// TIA Portal V20 export
// export: Created 2026-10-19T18:06:12.0545381Z, ExportSetting WithDefaults, DisplayName Totally Integrated Automation Portal, DisplayVersion V20 Update 6, DisplayName TIA Portal Openness, DisplayVersion V20 Update 6, DisplayName TIA Portal Version Control Interface, DisplayVersion V20 Update 6, DisplayName SINAMICS Startdrive Advanced, DisplayVersion V20 SP1, DisplayName SINAMICS Startdrive G130, G150, S120, S150, SINAMICS MV, G220, S200, S210, DisplayVersion V20 SP1, DisplayName SINAMICS Startdrive G110M, G120, G120C, G120D, G120P, G115D, DisplayVersion V20 SP1, DisplayName STEP 7 Professional, DisplayVersion V20 Update 6, DisplayName STEP 7 Safety, DisplayVersion V20 Update 2, DisplayName WinCC Basic/Comfort/Advanced, DisplayVersion V20 Update 6, DisplayName WinCC Unified, DisplayVersion V20 Update 6
FUNCTION "MT_ACT_Application" : Void   // FC30, LAD
{ S7_Optimized_Access := 'FALSE' }
VERSION : 0.1
// stored: AutoNumber true, IsIECCheckEnabled false, SetENOAutomatically false, UDAEnableTagReadback false
BEGIN

REGION Network 1: Cyclic Weighing Data
   // All the cyclical read and write commands can be issued from this Function Block.
   // The cyclic commands are triggered following a positive trigger. These commands are Tare Immediate, Tare Stable, Zero Immediate, Zero Stable, Pretare and Clear Tare. 
   // Upon successful execution of these commands, the DONE output bit will be set ON.
   // ERROR output bit will be set on if there is an error with the command execution.
   // Note: Only one cyclic command is possible at any one time.
   // If Net weight is required after executed a zero or tare command, insert decimal value "3" into the "WeightCmd" variable before triggering the cyclic scale command. Else, with decimal value "1" in the "WeightCmd" variable, the Function Block will return Gross Weight after the cyclic scale command. 
   // "DataOK" bit is set ON when the scale is in operation mode, not overloaded and not underload.
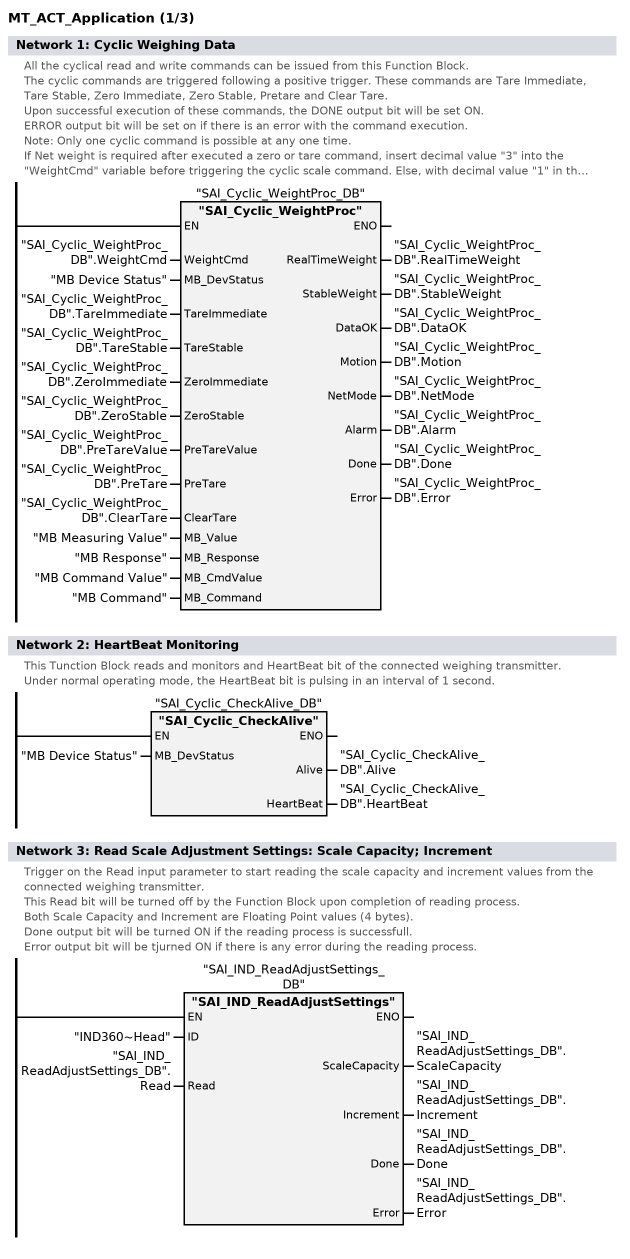
   RUNG wire#powerrail
      "SAI_Cyclic_WeightProc_DB"(WeightCmd := "SAI_Cyclic_WeightProc_DB".WeightCmd, MB_DevStatus := "MB Device Status", TareImmediate := "SAI_Cyclic_WeightProc_DB".TareImmediate, TareStable := "SAI_Cyclic_WeightProc_DB".TareStable, ZeroImmediate := "SAI_Cyclic_WeightProc_DB".ZeroImmediate, ZeroStable := "SAI_Cyclic_WeightProc_DB".ZeroStable, PreTareValue := "SAI_Cyclic_WeightProc_DB".PreTareValue, PreTare := "SAI_Cyclic_WeightProc_DB".PreTare, ClearTare := "SAI_Cyclic_WeightProc_DB".ClearTare, MB_Value := "MB Measuring Value", MB_Response := "MB Response", MB_CmdValue := "MB Command Value", MB_Command := "MB Command", RealTimeWeight => "SAI_Cyclic_WeightProc_DB".RealTimeWeight, StableWeight => "SAI_Cyclic_WeightProc_DB".StableWeight, DataOK => "SAI_Cyclic_WeightProc_DB".DataOK, Motion => "SAI_Cyclic_WeightProc_DB".Motion, NetMode => "SAI_Cyclic_WeightProc_DB".NetMode, Alarm => "SAI_Cyclic_WeightProc_DB".Alarm, Done => "SAI_Cyclic_WeightProc_DB".Done, Error => "SAI_Cyclic_WeightProc_DB".Error)
   END_RUNG
   // the same network as SCL:
   "SAI_Cyclic_WeightProc_DB"(WeightCmd := "SAI_Cyclic_WeightProc_DB".WeightCmd,   // "SAI_Cyclic_WeightProc"
                           MB_DevStatus := "MB Device Status",
                           TareImmediate := "SAI_Cyclic_WeightProc_DB".TareImmediate,
                           TareStable := "SAI_Cyclic_WeightProc_DB".TareStable,
                           ZeroImmediate := "SAI_Cyclic_WeightProc_DB".ZeroImmediate,
                           ZeroStable := "SAI_Cyclic_WeightProc_DB".ZeroStable,
                           PreTareValue := "SAI_Cyclic_WeightProc_DB".PreTareValue,
                           PreTare := "SAI_Cyclic_WeightProc_DB".PreTare,
                           ClearTare := "SAI_Cyclic_WeightProc_DB".ClearTare,
                           MB_Value := "MB Measuring Value",
                           MB_Response := "MB Response",
                           MB_CmdValue := "MB Command Value",
                           MB_Command := "MB Command",
                           RealTimeWeight => "SAI_Cyclic_WeightProc_DB".RealTimeWeight,
                           StableWeight => "SAI_Cyclic_WeightProc_DB".StableWeight,
                           DataOK => "SAI_Cyclic_WeightProc_DB".DataOK,
                           Motion => "SAI_Cyclic_WeightProc_DB".Motion,
                           NetMode => "SAI_Cyclic_WeightProc_DB".NetMode,
                           Alarm => "SAI_Cyclic_WeightProc_DB".Alarm,
                           Done => "SAI_Cyclic_WeightProc_DB".Done,
                           Error => "SAI_Cyclic_WeightProc_DB".Error);
END_REGION

REGION Network 2: HeartBeat Monitoring
   // This Tunction Block reads and monitors and HeartBeat bit of the connected weighing transmitter.
   // Under normal operating mode, the HeartBeat bit is pulsing in an interval of 1 second.
   RUNG wire#powerrail
      "SAI_Cyclic_CheckAlive_DB"(MB_DevStatus := "MB Device Status", Alive => "SAI_Cyclic_CheckAlive_DB".Alive, HeartBeat => "SAI_Cyclic_CheckAlive_DB".HeartBeat)
   END_RUNG
   // the same network as SCL:
   "SAI_Cyclic_CheckAlive_DB"(MB_DevStatus := "MB Device Status",   // "SAI_Cyclic_CheckAlive"
                           Alive => "SAI_Cyclic_CheckAlive_DB".Alive,
                           HeartBeat => "SAI_Cyclic_CheckAlive_DB".HeartBeat);
END_REGION

REGION Network 3: Read Scale Adjustment Settings: Scale Capacity; Increment
   // Trigger on the Read input parameter to start reading the scale capacity and increment values from the connected weighing transmitter.
   // This Read bit will be turned off by the Function Block upon completion of reading process.
   // Both Scale Capacity and Increment are Floating Point values (4 bytes).
   // Done output bit will be turned ON if the reading process is successfull.
   // Error output bit will be tjurned ON if there is any error during the reading process.
   RUNG wire#powerrail
      "SAI_IND_ReadAdjustSettings_DB"(ID := "IND360~Head", Read := "SAI_IND_ReadAdjustSettings_DB".Read, ScaleCapacity => "SAI_IND_ReadAdjustSettings_DB".ScaleCapacity, Increment => "SAI_IND_ReadAdjustSettings_DB".Increment, Done => "SAI_IND_ReadAdjustSettings_DB".Done, Error => "SAI_IND_ReadAdjustSettings_DB".Error)
   END_RUNG
   // the same network as SCL:
   "SAI_IND_ReadAdjustSettings_DB"(ID := "IND360~Head",   // "SAI_IND_ReadAdjustSettings"
                           Read := "SAI_IND_ReadAdjustSettings_DB".Read,
                           ScaleCapacity => "SAI_IND_ReadAdjustSettings_DB".ScaleCapacity,
                           Increment => "SAI_IND_ReadAdjustSettings_DB".Increment,
                           Done => "SAI_IND_ReadAdjustSettings_DB".Done,
                           Error => "SAI_IND_ReadAdjustSettings_DB".Error);
END_REGION

REGION Network 4: Write new Scale Adjustment Settings: Scale Capacity; Increment
   // Trigger on the Write input parameter to start writing the new scale capacity and increment settings to the connected weighing transmitter.
   // Both Scale Capacity and Increment are Floating Point values (4 bytes).
   // Make sure both settings are valid and correct before triggering the Write input bit.
   // This Write bit will be turned off by the Function Block upon completion of writing process.
   // Done output bit will be set ON if the reading process is successfull.
   // Error output bit will be set ON if there is any error during the reading process.
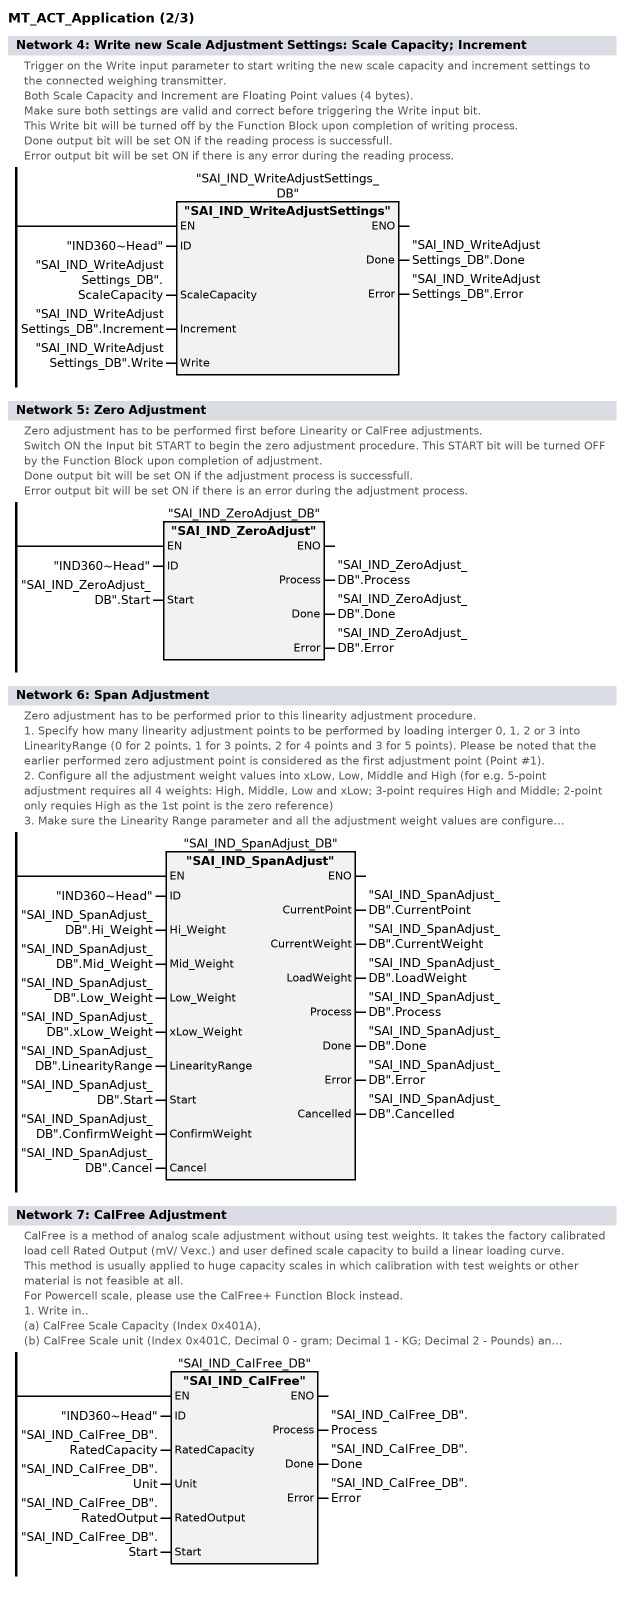
   RUNG wire#powerrail
      "SAI_IND_WriteAdjustSettings_DB"(ID := "IND360~Head", ScaleCapacity := "SAI_IND_WriteAdjustSettings_DB".ScaleCapacity, Increment := "SAI_IND_WriteAdjustSettings_DB".Increment, Write := "SAI_IND_WriteAdjustSettings_DB".Write, Done => "SAI_IND_WriteAdjustSettings_DB".Done, Error => "SAI_IND_WriteAdjustSettings_DB".Error)
   END_RUNG
   // the same network as SCL:
   "SAI_IND_WriteAdjustSettings_DB"(ID := "IND360~Head",   // "SAI_IND_WriteAdjustSettings"
                           ScaleCapacity := "SAI_IND_WriteAdjustSettings_DB".ScaleCapacity,
                           Increment := "SAI_IND_WriteAdjustSettings_DB".Increment,
                           Write := "SAI_IND_WriteAdjustSettings_DB".Write,
                           Done => "SAI_IND_WriteAdjustSettings_DB".Done,
                           Error => "SAI_IND_WriteAdjustSettings_DB".Error);
END_REGION

REGION Network 5: Zero Adjustment
   // Zero adjustment has to be performed first before Linearity or CalFree adjustments.
   // Switch ON the Input bit START to begin the zero adjustment procedure. This START bit will be turned OFF by the Function Block upon completion of adjustment. 
   // Done output bit will be set ON if the adjustment process is successfull.
   // Error output bit will be set ON if there is an error during the adjustment process.
   RUNG wire#powerrail
      "SAI_IND_ZeroAdjust_DB"(ID := "IND360~Head", Start := "SAI_IND_ZeroAdjust_DB".Start, Process => "SAI_IND_ZeroAdjust_DB".Process, Done => "SAI_IND_ZeroAdjust_DB".Done, Error => "SAI_IND_ZeroAdjust_DB".Error)
   END_RUNG
   // the same network as SCL:
   "SAI_IND_ZeroAdjust_DB"(ID := "IND360~Head",   // "SAI_IND_ZeroAdjust"
                           Start := "SAI_IND_ZeroAdjust_DB".Start,
                           Process => "SAI_IND_ZeroAdjust_DB".Process,
                           Done => "SAI_IND_ZeroAdjust_DB".Done,
                           Error => "SAI_IND_ZeroAdjust_DB".Error);
END_REGION

REGION Network 6: Span Adjustment
   // Zero adjustment has to be performed prior to this linearity adjustment procedure.
   // 
   // 1. Specify how many linearity adjustment points to be performed by loading interger 0, 1, 2 or 3 into LinearityRange (0 for 2 points, 1 for 3 points, 2 for 4 points and 3 for 5 points). Please be noted that the earlier performed zero adjustment point is considered as the first adjustment point (Point #1).
   // 
   // 2. Configure all the adjustment weight values into xLow, Low, Middle and High (for e.g. 5-point adjustment requires all 4 weights: High, Middle, Low and xLow; 3-point requires High and Middle; 2-point only requies High as the 1st point is the zero reference)
   // 
   // 3. Make sure the Linearity Range parameter and all the adjustment weight values are configured correctly before starting the adjustment process. Invalid or incomplete parameters will cause the Function Block to turn on the Error output bit.
   // 
   // 4. Trigger ON  Input Start bit to start the span adjustment. This Start bit will be turned off by the Function Block upon completion/ cancellation or error condition. 
   // 
   // 5. Once started, CurrentPoint shows the current linearity point to be adjusted; CurrentWeight shows current adjustment weight to be loaded onto the scale. The LoadWeight output bit will be set ON to request for new adjustment weight. 
   // 
   // 6. After loading the new adjustment weight, acknowledge this by triggering the ConfirmWeight parameter (boolean) ON. The Function Block will then proceed to the next adjustment point and turn off this ConfirmWeight bit.
   // 
   // 7. Output bit - Process signifies that the adjustment of current point is in process.
   // 
   // 8. Input Parameter Bit Cancel is used to cancel/ abort the adjustment process
   RUNG wire#powerrail
      "SAI_IND_SpanAdjust_DB"(ID := "IND360~Head", Hi_Weight := "SAI_IND_SpanAdjust_DB".Hi_Weight, Mid_Weight := "SAI_IND_SpanAdjust_DB".Mid_Weight, Low_Weight := "SAI_IND_SpanAdjust_DB".Low_Weight, xLow_Weight := "SAI_IND_SpanAdjust_DB".xLow_Weight, LinearityRange := "SAI_IND_SpanAdjust_DB".LinearityRange, Start := "SAI_IND_SpanAdjust_DB".Start, ConfirmWeight := "SAI_IND_SpanAdjust_DB".ConfirmWeight, Cancel := "SAI_IND_SpanAdjust_DB".Cancel, CurrentPoint => "SAI_IND_SpanAdjust_DB".CurrentPoint, CurrentWeight => "SAI_IND_SpanAdjust_DB".CurrentWeight, LoadWeight => "SAI_IND_SpanAdjust_DB".LoadWeight, Process => "SAI_IND_SpanAdjust_DB".Process, Done => "SAI_IND_SpanAdjust_DB".Done, Error => "SAI_IND_SpanAdjust_DB".Error, Cancelled => "SAI_IND_SpanAdjust_DB".Cancelled)
   END_RUNG
   // the same network as SCL:
   "SAI_IND_SpanAdjust_DB"(ID := "IND360~Head",   // "SAI_IND_SpanAdjust"
                           Hi_Weight := "SAI_IND_SpanAdjust_DB".Hi_Weight,
                           Mid_Weight := "SAI_IND_SpanAdjust_DB".Mid_Weight,
                           Low_Weight := "SAI_IND_SpanAdjust_DB".Low_Weight,
                           xLow_Weight := "SAI_IND_SpanAdjust_DB".xLow_Weight,
                           LinearityRange := "SAI_IND_SpanAdjust_DB".LinearityRange,
                           Start := "SAI_IND_SpanAdjust_DB".Start,
                           ConfirmWeight := "SAI_IND_SpanAdjust_DB".ConfirmWeight,
                           Cancel := "SAI_IND_SpanAdjust_DB".Cancel,
                           CurrentPoint => "SAI_IND_SpanAdjust_DB".CurrentPoint,
                           CurrentWeight => "SAI_IND_SpanAdjust_DB".CurrentWeight,
                           LoadWeight => "SAI_IND_SpanAdjust_DB".LoadWeight,
                           Process => "SAI_IND_SpanAdjust_DB".Process,
                           Done => "SAI_IND_SpanAdjust_DB".Done,
                           Error => "SAI_IND_SpanAdjust_DB".Error,
                           Cancelled => "SAI_IND_SpanAdjust_DB".Cancelled);
END_REGION

REGION Network 7: CalFree Adjustment
   // CalFree is a method of analog scale adjustment without using test weights. It takes the factory calibrated load cell Rated Output (mV/ Vexc.) and user defined scale capacity to build a linear loading curve.
   // This method is usually applied to huge capacity scales in which calibration with test weights or other material is not feasible at all. 
   // 
   // For Powercell scale, please use the CalFree+ Function Block instead.
   // 
   // 1. Write in.. 
   // (a) CalFree Scale Capacity (Index 0x401A), 
   // (b) CalFree Scale unit (Index 0x401C, Decimal 0 - gram; Decimal 1 - KG; Decimal 2 - Pounds) and 
   // (c) Load Cells' averaged Rated Output (Index 0x401D, in mV/V)
   // **Make sure the transmitter's scale capacity has already been configured to the same value as CalFree Capacity prior to this CalFree adjustment.
   // 
   // 2. Trigger Input bit Start for CalFree adjustment (Index 0x401A)
   // 
   // 3. Output bit Done will be turned ON after successful completion of the process
   // Error output bit will be turned ON if there is an error during the adjustment process
   RUNG wire#powerrail
      "SAI_IND_CalFree_DB"(ID := "IND360~Head", RatedCapacity := "SAI_IND_CalFree_DB".RatedCapacity, Unit := "SAI_IND_CalFree_DB".Unit, RatedOutput := "SAI_IND_CalFree_DB".RatedOutput, Start := "SAI_IND_CalFree_DB".Start, Process => "SAI_IND_CalFree_DB".Process, Done => "SAI_IND_CalFree_DB".Done, Error => "SAI_IND_CalFree_DB".Error)
   END_RUNG
   // the same network as SCL:
   "SAI_IND_CalFree_DB"(ID := "IND360~Head",   // "SAI_IND_CalFree"
                        RatedCapacity := "SAI_IND_CalFree_DB".RatedCapacity,
                        Unit := "SAI_IND_CalFree_DB".Unit,
                        RatedOutput := "SAI_IND_CalFree_DB".RatedOutput,
                        Start := "SAI_IND_CalFree_DB".Start,
                        Process => "SAI_IND_CalFree_DB".Process,
                        Done => "SAI_IND_CalFree_DB".Done,
                        Error => "SAI_IND_CalFree_DB".Error);
END_REGION

REGION Network 8: Alibi Record Read
   // Use this Function Block to read one alibi record. 
   // 1. Set the alibi transaction number to be read.
   // 2. Toggle the Get_Record bit to perform read. Alibi record will be written into Alibi_Array (an array of 44 Bytes).  
   // 3. The read alibi record transaction gross, net and tare weights (all LREAL format) as well as weight unit are available at the FB's output.
   // 4. the Alibi_Array structure data format is as below:
   // 
   // For Base, RateControl, Tank Vessel:
   // Struct(44 Bytes)
   // {
   // Byte[20]: Date & time; //ASCII String  =>Byte0-19
   // Long:     Transaction Number;            =>Byte20-23
   // Float32:  Gross Weight;                       =>Byte24-27
   // Float32:  Net Weight;                           =>Byte28-31
   // Float32:  Tare Weight;                         =>Byte32-35
   // Byte:     Tare Mode;                              =>Byte36
   // Byte:     Unit;                                          =>Byte37
   // Byte[6]:  Not Used;                              =>Byte38-43
   // }
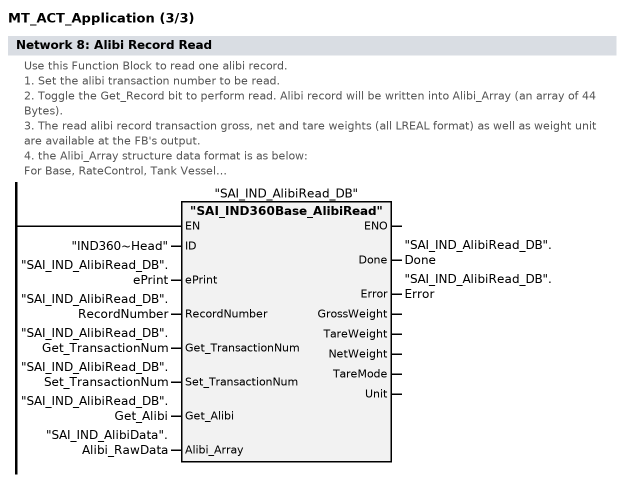
   RUNG wire#powerrail
      "SAI_IND_AlibiRead_DB"(ID := "IND360~Head", ePrint := "SAI_IND_AlibiRead_DB".ePrint, RecordNumber := "SAI_IND_AlibiRead_DB".RecordNumber, Get_TransactionNum := "SAI_IND_AlibiRead_DB".Get_TransactionNum, Set_TransactionNum := "SAI_IND_AlibiRead_DB".Set_TransactionNum, Get_Alibi := "SAI_IND_AlibiRead_DB".Get_Alibi, Alibi_Array := "SAI_IND_AlibiData".Alibi_RawData, Done => "SAI_IND_AlibiRead_DB".Done, Error => "SAI_IND_AlibiRead_DB".Error, GrossWeight =>, TareWeight =>, NetWeight =>, TareMode =>, Unit =>)
   END_RUNG
   // the same network as SCL:
   "SAI_IND_AlibiRead_DB"(ID := "IND360~Head",   // "SAI_IND360Base_AlibiRead"
                          ePrint := "SAI_IND_AlibiRead_DB".ePrint,
                          RecordNumber := "SAI_IND_AlibiRead_DB".RecordNumber,
                          Get_TransactionNum := "SAI_IND_AlibiRead_DB".Get_TransactionNum,
                          Set_TransactionNum := "SAI_IND_AlibiRead_DB".Set_TransactionNum,
                          Get_Alibi := "SAI_IND_AlibiRead_DB".Get_Alibi,
                          Alibi_Array := "SAI_IND_AlibiData".Alibi_RawData,
                          Done => "SAI_IND_AlibiRead_DB".Done,
                          Error => "SAI_IND_AlibiRead_DB".Error);
END_REGION
END_FUNCTION
